{attribute 'qualified_only' := ''}
{attribute 'strict' := ''}
TYPE E_TrackType :
(
	TRACKTYPE_NONE := 0,
	TRACKTYPE_FERRY := 1,
	TRACKTYPE_LINE := 2,
	TRACKTYPE_CIRCLE := 3,
	TRACKTYPE_FORK := 4
);
END_TYPE

(* stored: Version 1.1.0.1, ProductVersion 3.1.4024.12
   DUT E_TrackType: Id {c703414d-e36d-4087-91c6-679bb3713735} *)
